// TIA Portal V20 export
// export: Created 2026-10-20T12:53:57.0288295Z, ExportSetting WithDefaults, DisplayName Totally Integrated Automation Portal, DisplayVersion V20 Update 6, DisplayName TIA Portal Openness, DisplayVersion V20 Update 6, DisplayName TIA Portal Version Control Interface, DisplayVersion V20 Update 6, DisplayName SINAMICS Startdrive Advanced, DisplayVersion V20 SP1, DisplayName SINAMICS Startdrive G130, G150, S120, S150, SINAMICS MV, G220, S200, S210, DisplayVersion V20 SP1, DisplayName SINAMICS Startdrive G110M, G120, G120C, G120D, G120P, G115D, DisplayVersion V20 SP1, DisplayName STEP 7 Professional, DisplayVersion V20 Update 6, DisplayName STEP 7 Safety, DisplayVersion V20 Update 2, DisplayName WinCC Basic/Comfort/Advanced, DisplayVersion V20 Update 6, DisplayName WinCC Unified, DisplayVersion V20 Update 6
FUNCTION "VTD_Order_FC" : Void   // FC45, SCL
{ S7_Optimized_Access := 'TRUE' }
VERSION : 0.1
// stored: AutoNumber true, IsIECCheckEnabled false, SetENOAutomatically false, UDAEnableTagReadback false
   VAR_INPUT
      i_Sys : UInt;
      Level : UInt;
   END_VAR
   VAR_IN_OUT
      StepTable_0 : "OrderTable_UDT";
   END_VAR
   VAR_TEMP
      StrSys : String;
      Concat1 : String;
      StrLev : String;
      Concat2 : String;
      ID : DInt;
   END_VAR
BEGIN
   #StrSys := UINT_TO_STRING(#i_Sys);
   // Remove "+"
   IF #StrSys[1] = '+' THEN
       #StrSys := RIGHT(IN := #StrSys, L := LEN(#StrSys) - 1);
   END_IF;

   #StrLev := UINT_TO_STRING(#Level);

   // Remove "+"
   IF #StrLev[1] = '+' THEN
       #StrLev := RIGHT(IN := #StrLev, L := LEN(#StrLev) - 1);
   END_IF;

   // Build ID
   #Concat1 := CONCAT(IN1 := '300', IN2 := #StrLev);
   #Concat2 := CONCAT(IN1 := #Concat1, IN2 := '0');
   #ID := STRING_TO_DINT(IN := CONCAT(IN1 := #Concat2, IN2 := #StrSys));

   "Feed_Steptable_FC"(CurrentTime := "Time".CurrentLocalTime,
                       Task_Type := 1,
                       Source_Location := 0,
                       Destination_Location := #ID,
                       Pallet_Type := 'C',
                       Pallet_Alignment := 'N',
                       Shuttle_ID:=0,
                       StepTable := #"StepTable_0");
END_FUNCTION
